// TIA Portal V20 export
Screen "Pop-up_SPEC_FUNCTIONS_Popup"  530x171
  ScreenItem "Background" at 0,0 size 532x171  Type=HmiRectangle
  ScreenItem "Overview_Special" at 1,1 size 523x25  Type=HmiTextBox
  ScreenItem "Cancel Mode" at 408,-3 size 116x58  Type=HmiButton
  ScreenItem "Stop Mode" at 10,38 size 90x60  Type=HmiButton
  ScreenItem "Mode Home Position" at 10,101 size 90x60  Type=HmiButton
  ScreenItem "Mode End of Cycle" at 103,38 size 90x60  Type=HmiButton
  ScreenItem "Mode Release Enty" at 103,101 size 90x60  Type=HmiButton
  ScreenItem "Mode Single Step" at 196,38 size 90x60  Type=HmiButton
  ScreenItem "Mode SingleStep plus1" at 196,101 size 90x60  Type=HmiButton
  ScreenItem "Mode Empty Position" at 289,38 size 90x60  Type=HmiButton
  ScreenItem "Mode WithoutPart Dryrun" at 289,101 size 90x60  Type=HmiButton
  ScreenItem "Textfield_SelectedOPMode" at 196,1 size 34x24  Type=HmiTextBox
  ScreenItem "stop_Foreground_Blocked" at 10,38 size 90x60  Type=HmiGraphicView
  ScreenItem "stop_Blocked" at 13,43 size 14x14  Type=HmiGraphicView
  ScreenItem "home_Foreground_Blocked" at 11,101 size 90x60  Type=HmiGraphicView
  ScreenItem "home_Blocked" at 13,103 size 14x14  Type=HmiGraphicView
  ScreenItem "eoc_Foreground_Blocked" at 103,38 size 90x60  Type=HmiGraphicView
  ScreenItem "eoc_Blocked" at 105,43 size 14x14  Type=HmiGraphicView
  ScreenItem "relEntry_Foreground_Blocked" at 103,101 size 90x60  Type=HmiGraphicView
  ScreenItem "relEntry_Blocked" at 104,103 size 14x14  Type=HmiGraphicView
  ScreenItem "singleStep_Foreground_Blocked" at 196,38 size 90x60  Type=HmiGraphicView
  ScreenItem "singleStep_Blocked" at 197,43 size 14x14  Type=HmiGraphicView
  ScreenItem "stepPlus_Foreground_Blocked" at 196,101 size 90x60  Type=HmiGraphicView
  ScreenItem "stepPlus_Blocked" at 198,103 size 14x14  Type=HmiGraphicView
  ScreenItem "emptyLine_Foreground_Blocked" at 289,37 size 90x60  Type=HmiGraphicView
  ScreenItem "emptyLine_Blocked" at 293,43 size 14x14  Type=HmiGraphicView
  ScreenItem "noPart_Foreground_Blocked" at 289,101 size 90x60  Type=HmiGraphicView
  ScreenItem "noPart_Blocked" at 292,103 size 14x14  Type=HmiGraphicView
  ScreenItem "Button_1" at 408,103 size 116x58  Type=HmiButton
